{region 'Documentation'}
(*!
<summary>Checks that the rising-edge count is greater than the strict limit.</summary>
<description>

Observation and accumulated-count handling come from AssertionEdgeCountBase. Evaluate
checks the held count independently of Enable; reset clears the count and baseline.

</description>
*)
{endregion}
FUNCTION_BLOCK AssertRisingEdgeCntGreaterThan EXTENDS AssertionEdgeCountBase
VAR_INPUT
    Minimum : UINT; //! Exclusive lower bound; the actual value or count must be greater.
END_VAR

SUPER^();

{region 'Documentation'}
(*!
<summary>Observe through the base, then evaluate the count with Error priority.</summary>
*)
{endregion}
METHOD PROTECTED Assert
VAR
    Message : STRING(GVL_Constants.MessageLength);
    MinimumText : STRING(GVL_Constants.AssertionValueLength);
    ActualText : STRING(GVL_Constants.AssertionValueLength);
END_VAR
SUPER^.Assert();

IF NOT EvaluationActive THEN
    RETURN;
END_IF;

IF Result = E_Result.Error THEN
    RETURN;
END_IF;

IF Result = E_Result.Failed THEN
    RETURN;
END_IF;

IF EdgeCount <= Minimum THEN
    MinimumText := UINT_TO_STRING(Minimum);
    ActualText := UINT_TO_STRING(EdgeCount);
    Message := CONCAT('Assertion failed: rising edge count is not greater than limit. Minimum = ',
        MinimumText);
    Message := CONCAT(Message, ', Actual = ');
    Message := CONCAT(Message, ActualText);
    Message := CONCAT(Message, '.');
    Fail(Message := Message);
    RETURN;
END_IF;

Pass();
END_METHOD

{region 'Documentation'}
(*!
<summary>Recognize a rising edge without changing observation state.</summary>
*)
{endregion}
METHOD PROTECTED IsMatchingEdge : BOOL //! TRUE when PreviousValue and CurrentValue form the edge selected by this Assertion.
VAR_INPUT
    PreviousValue : BOOL; //! Signal value from the preceding active observation.
    CurrentValue : BOOL; //! Signal value from the current active observation.
END_VAR
IsMatchingEdge := NOT PreviousValue AND CurrentValue;
END_METHOD

END_FUNCTION_BLOCK

(* stored: Version 1.1.0.1
   POU AssertRisingEdgeCntGreaterThan: Id {8129a732-d2fe-484b-828e-3e6bc4cc3ecd}, SpecialFunc None
   Folder Internal: Id {9bd8db1c-4c00-4fde-bf6e-964a91ad72ae}
   Method Assert: Id {153fdcfb-16d9-4e6c-aea2-d4b6682c839f}
   Method IsMatchingEdge: Id {bf9445c4-8640-4b52-91fa-83798b8e381b} *)
